(*
SPDX-FileCopyrightText: © 2026 Oleksandr Tiutyk <trofimich@gmail.com>
SPDX-License-Identifier: MIT
License: https://opensource.org/license/mit
*)

(*!
<summary>
Beckhoff EL1502: 2-channel up/down counter terminal (24 V DC, 100 kHz).
</summary>
<description>
Requires the 2Ch. Counter assignment: TxPDOs 0x1A00/0x1A01 and RxPDOs 0x1600/0x1601.
Each channel is a 32-bit counter with 16-bit status/control; direction is configured through CoE.
The factory 1Ch. +/- Counter assignment 0x1A02/0x1602 is not represented.
This model does not provide two independent hardware up/down input pairs.
When used for I/O, link located fields or their containing buffers to the matching selected PDOs.
The record is not a packed wire buffer; compiler padding is not part of the device specification.
Unlinked/default values do not prove valid I/O. The caller evaluates bus/channel validity before use.
Use one owner task per instance and externally synchronize other access; multi-field snapshots are not atomic.
Copies store data without creating hardware links. Keep borrowed field references valid while consumers are bound.
This passive record performs no validation, synchronization, configuration or protocol advancement.
</description>
*)
TYPE EL1502 :
STRUCT
	Ch1 : COUNTER_CHANNEL;
	Ch2 : COUNTER_CHANNEL;
END_STRUCT
END_TYPE

(* stored: Version 1.1.0.1, ProductVersion 3.1.4026.20
   DUT EL1502: Id {00e1875c-2a7c-42d9-b25d-e52955f667dd} *)
